FUNCTION_BLOCK basicMotorGenerico (* Logica unica do motor generico (partida direta ou inversor) *)
  (* Standard: 61499-2 *)
  (* Version 2.2, 12/11/2026, Hidryco, Hidryco, 2.2: cfgFalhaNA (contato de falha NA, dosagem 800). 2.1: raio do gerador vermelho (3) so com a carga liberada, a planta nos geradores E o motor ligado (igual ao Motor_VS, gradeamento e UV); liberado e parado = cinza (2). 2.0: velocidade da IHM/SCADA (stsVelocidadeIhm, antes stsVelocidadeHz) em %%: com inversor = fldVelocidadePct (LSP 0 %% a HSP 100 %%), sem inversor = 0 ou 100 %%; referencia e manual continuam em Hz. 1.9: velocidade manual (stpVelocidadeManual) em Hz; saidas stsVelocidadeHz/stsReferenciaHz para a IHM (conversao no CLP, 60 Hz = 100 %). 1.8: IHM: velocidade e referencia no maximo 1 vez por segundo com o motor ligado (antes a cada 0,1 %); o plug/processo (CNF_SPEED) continua na hora. 1.7: saida stsFalhaAtiva (falha presente agora: emergencia, termica, acionamento ou comunicacao) no CNF_HMI. 1.6: protecao termica nao memoriza - sai sozinha quando normaliza (sem reset). 1.5: reset so libera a falha de parada com o motor parado (antes liberava com o motor ainda ligado e a supervisao nao recomecava). 1.1: refeito no padrao SE.App2CommonProcess - eventos por grupo de dados, saidas so na mudanca, supervisao por E_DELAY (MON_T/MON_RESET/MON_MAX), horimetro e partidas pelo devMntCalc, escala linear com limites. 1.4: horimetro proprio com resolucao de 1 s (E_CYCLE + PERSISTENCE), termica NF por padrao *)
  PACKAGE Hidryco.HidrycoLib;
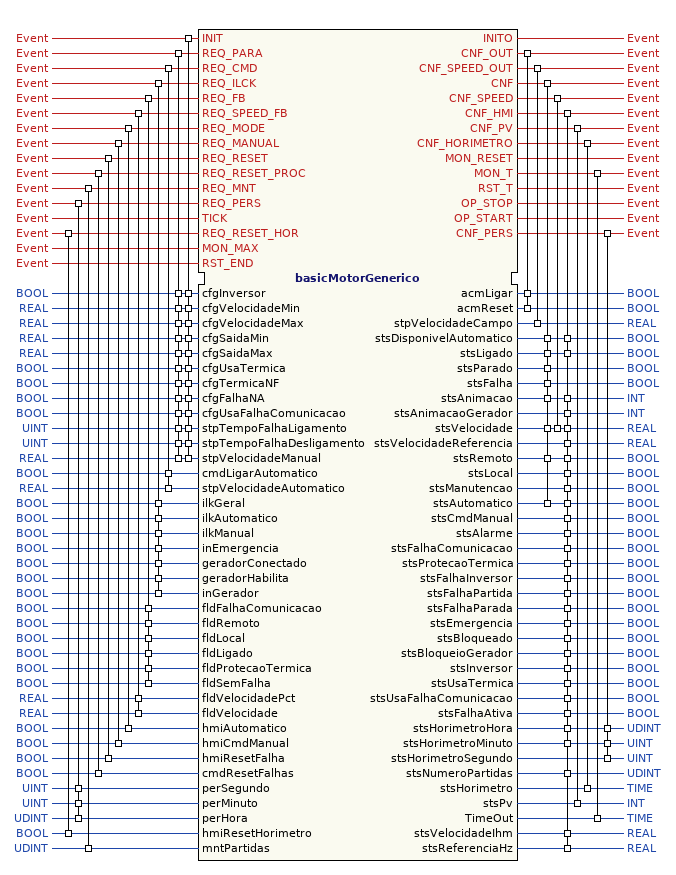
  EVENT_INPUT
    INIT WITH cfgInversor, cfgVelocidadeMin, cfgVelocidadeMax, cfgSaidaMin, cfgSaidaMax, cfgUsaTermica, cfgTermicaNF, cfgFalhaNA, cfgUsaFalhaComunicacao, stpTempoFalhaLigamento, stpTempoFalhaDesligamento, stpVelocidadeManual; (* Inicializacao (configuracao da instancia) *)
    REQ_PARA WITH cfgInversor, cfgVelocidadeMin, cfgVelocidadeMax, cfgSaidaMin, cfgSaidaMax, cfgUsaTermica, cfgTermicaNF, cfgFalhaNA, cfgUsaFalhaComunicacao, stpTempoFalhaLigamento, stpTempoFalhaDesligamento, stpVelocidadeManual; (* Atualizacao de parametros (IHM) *)
    REQ_CMD WITH cmdLigarAutomatico, stpVelocidadeAutomatico; (* Comando e referencia do processo *)
    REQ_ILCK WITH ilkGeral, ilkAutomatico, ilkManual, inEmergencia, geradorConectado, geradorHabilita, inGerador; (* Intertravamentos, emergencia e gerador *)
    REQ_FB WITH fldFalhaComunicacao, fldRemoto, fldLocal, fldLigado, fldProtecaoTermica, fldSemFalha; (* Sinais de campo *)
    REQ_SPEED_FB WITH fldVelocidade, fldVelocidadePct; (* Velocidade real do inversor *)
    REQ_MODE WITH hmiAutomatico; (* Modo automatico/manual (IHM) *)
    REQ_MANUAL WITH hmiCmdManual; (* Liga/desliga manual (IHM) *)
    REQ_RESET WITH hmiResetFalha; (* Reset de falhas (IHM) *)
    REQ_RESET_PROC WITH cmdResetFalhas; (* Reset de falhas (processo) *)
    REQ_MNT WITH mntPartidas; (* Numero de partidas do devMntCalc *)
    REQ_PERS WITH perSegundo, perMinuto, perHora; (* Horimetro lido do PERSISTENCE (READCNF) *)
    TICK; (* 1 s do E_CYCLE (so com o motor ligado) *)
    REQ_RESET_HOR WITH hmiResetHorimetro; (* Zera o horimetro (IHM) *)
    MON_MAX; (* Tempo de supervisao de partida/parada esgotado (E_DELAY) *)
    RST_END; (* Fim do pulso de reset (E_DELAY) *)
  END_EVENT
  EVENT_OUTPUT
    INITO; (* Inicializacao concluida *)
    CNF_OUT WITH acmLigar, acmReset; (* Saidas digitais de campo (na mudanca) *)
    CNF_SPEED_OUT WITH stpVelocidadeCampo; (* Referencia de velocidade para o campo (na mudanca) *)
    CNF WITH stsDisponivelAutomatico, stsLigado, stsParado, stsFalha, stsAnimacao, stsVelocidade, stsRemoto, stsAutomatico; (* Status para o processo (na mudanca) *)
    CNF_SPEED WITH stsVelocidade; (* Velocidade real (mudanca maior ou igual a 0,1 %) *)
    CNF_HMI WITH stsRemoto, stsLocal, stsManutencao, stsLigado, stsAutomatico, stsCmdManual, stsAnimacao, stsAnimacaoGerador, stsAlarme, stsFalhaComunicacao, stsProtecaoTermica, stsFalhaInversor, stsFalhaPartida, stsFalhaParada, stsEmergencia, stsBloqueado, stsBloqueioGerador, stsDisponivelAutomatico, stsVelocidade, stsVelocidadeReferencia, stsHorimetroHora, stsHorimetroMinuto, stsNumeroPartidas, stsInversor, stsUsaTermica, stsUsaFalhaComunicacao, stsFalhaAtiva, stsVelocidadeIhm, stsReferenciaHz; (* Status para a IHM (na mudanca) *)
    CNF_PV WITH stsPv; (* Estado ligado/parado para o devMntCalc (na mudanca) *)
    CNF_HORIMETRO WITH stsHorimetro; (* Tempo de operacao (na mudanca) *)
    MON_RESET; (* Cancela o tempo de supervisao (E_DELAY.STOP) - sai antes do MON_T *)
    MON_T WITH TimeOut; (* Inicia o tempo de supervisao (E_DELAY.START) *)
    RST_T; (* Inicia o pulso de reset (E_DELAY.START) *)
    OP_STOP; (* Para o E_CYCLE do horimetro - sai antes do OP_START *)
    OP_START; (* Inicia o E_CYCLE de 1 s do horimetro *)
    CNF_PERS WITH stsHorimetroSegundo, stsHorimetroMinuto, stsHorimetroHora; (* Grava o horimetro no PERSISTENCE (a cada minuto, na parada e no reset) *)
  END_EVENT
  VAR_INPUT
    cfgInversor : BOOL := FALSE; (* TRUE = motor com inversor (referencia de velocidade e medicoes) *)
    cfgVelocidadeMin : REAL := 0.0; (* Limite minimo da referencia de velocidade (%) *)
    cfgVelocidadeMax : REAL := 100.0; (* Limite maximo da referencia de velocidade (%) *)
    cfgSaidaMin : REAL := 0.0; (* Valor de campo equivalente a 0 % (referencia e realimentacao) *)
    cfgSaidaMax : REAL := 100.0; (* Valor de campo equivalente a 100 % (ex.: 100 = %, 60 = Hz, 10000 = Sulzer 0,01 %) *)
    cfgUsaTermica : BOOL := TRUE; (* TRUE = supervisiona a protecao termica *)
    cfgTermicaNF : BOOL := TRUE; (* TRUE = termica NF (FALSE no campo = atuada). Padrao NF (definido pelo usuario) *)
    cfgFalhaNA : BOOL := FALSE; (* TRUE = contato de falha do acionamento NA (TRUE no campo = falha, ligado em stsSemFalha). Padrao FALSE = NF (SEM FALHA) *)
    cfgUsaFalhaComunicacao : BOOL := TRUE; (* TRUE = considera o bit de falha de comunicacao da remota *)
    stpTempoFalhaLigamento : UINT; (* Tempo maximo para confirmar a partida (s). 0 = sem supervisao *)
    stpTempoFalhaDesligamento : UINT; (* Tempo maximo para confirmar a parada (s). 0 = sem supervisao *)
    stpVelocidadeManual : REAL; (* IHM: velocidade em manual em Hz (60 Hz = 100 %) *)
    cmdLigarAutomatico : BOOL; (* Comando ligar do processo (modo automatico) *)
    stpVelocidadeAutomatico : REAL; (* Referencia de velocidade do processo (%) *)
    ilkGeral : BOOL; (* Intertravamento geral (automatico e manual) *)
    ilkAutomatico : BOOL; (* Intertravamento so do automatico *)
    ilkManual : BOOL; (* Intertravamento so do manual *)
    inEmergencia : BOOL; (* Emergencia (TRUE = acionada): retira o comando e exige reset *)
    geradorConectado : BOOL; (* TRUE = o gerador pode alimentar este equipamento *)
    geradorHabilita : BOOL; (* Selecao do operador no CAT Gerador (HAB_GERADOR_EQUIP_n) *)
    inGerador : BOOL; (* TRUE = planta alimentada pelo gerador *)
    fldFalhaComunicacao : BOOL; (* Campo: falha de comunicacao da remota *)
    fldRemoto : BOOL; (* Campo: chave em remoto *)
    fldLocal : BOOL; (* Campo: chave em local *)
    fldLigado : BOOL; (* Campo: confirmacao de ligado *)
    fldProtecaoTermica : BOOL; (* Campo: protecao termica (ver cfgTermicaNF) *)
    fldSemFalha : BOOL; (* Campo: falha NF (TRUE = sem falha) *)
    fldVelocidadePct : REAL; (* Campo: velocidade do inversor em % (0 % no LSP, 100 % no HSP), so para a IHM *)
    fldVelocidade : REAL; (* Campo: velocidade real na unidade de cfgSaidaMin..cfgSaidaMax *)
    hmiAutomatico : BOOL; (* IHM: TRUE = automatico *)
    hmiCmdManual : BOOL; (* IHM: TRUE = ligar, FALSE = desligar (manual) *)
    hmiResetFalha : BOOL; (* IHM: reset de falhas (vale com TRUE) *)
    cmdResetFalhas : BOOL; (* Processo: reset de falhas (vale com TRUE) *)
    perSegundo : UINT; (* Horimetro persistido: segundos *)
    perMinuto : UINT; (* Horimetro persistido: minutos *)
    perHora : UDINT; (* Horimetro persistido: horas *)
    hmiResetHorimetro : BOOL; (* IHM: zera o horimetro (vale com TRUE) *)
    mntPartidas : UDINT; (* devMntCalc: numero de partidas *)
  END_VAR
  VAR_OUTPUT
    acmLigar : BOOL; (* Campo: comando liga *)
    acmReset : BOOL; (* Campo: pulso de reset (inversor/rele) *)
    stpVelocidadeCampo : REAL; (* Campo: referencia de velocidade (cfgSaidaMin..cfgSaidaMax) *)
    stsDisponivelAutomatico : BOOL; (* Pode ser comandado pelo automatico agora *)
    stsLigado : BOOL; (* Motor ligado (confirmacao de campo) *)
    stsParado : BOOL; (* Motor parado *)
    stsFalha : BOOL; (* Alguma falha memorizada (exige reset) *)
    stsAnimacao : INT; (* 0 desligado, 1 ligado, 2 falha, 3 manutencao *)
    stsAnimacaoGerador : INT; (* 0 nao conectado, 1 conectado, 2 selecionado, 3 selecionado e gerador ligado *)
    stsVelocidade : REAL; (* Velocidade real (%); partida direta: 0 ou 100 *)
    stsVelocidadeReferencia : REAL; (* Referencia de velocidade em uso (%) *)
    stsRemoto : BOOL; (* Chave em remoto *)
    stsLocal : BOOL; (* Chave em local *)
    stsManutencao : BOOL; (* Chave na posicao 0 *)
    stsAutomatico : BOOL; (* Modo automatico *)
    stsCmdManual : BOOL; (* Comando manual em vigor *)
    stsAlarme : BOOL; (* Falha memorizada ou falha de comunicacao *)
    stsFalhaComunicacao : BOOL; (* Falha de comunicacao *)
    stsProtecaoTermica : BOOL; (* Termica memorizada *)
    stsFalhaInversor : BOOL; (* Falha do acionamento memorizada *)
    stsFalhaPartida : BOOL; (* Nao confirmou partida no tempo *)
    stsFalhaParada : BOOL; (* Nao confirmou parada no tempo *)
    stsEmergencia : BOOL; (* Emergencia memorizada *)
    stsBloqueado : BOOL; (* Intertravamento ativo no modo atual *)
    stsBloqueioGerador : BOOL; (* Bloqueado pelo gerador *)
    stsInversor : BOOL; (* Copia de cfgInversor (IHM) *)
    stsUsaTermica : BOOL; (* Copia de cfgUsaTermica (IHM) *)
    stsUsaFalhaComunicacao : BOOL; (* Copia de cfgUsaFalhaComunicacao (IHM) *)
    stsFalhaAtiva : BOOL; (* Falha ativa (agora, sem memoria): emergencia, termica, acionamento ou comunicacao *)
    stsHorimetroHora : UDINT; (* Horimetro (h) *)
    stsHorimetroMinuto : UINT; (* Horimetro (min, 0-59) *)
    stsHorimetroSegundo : UINT; (* Horimetro (s, 0-59) *)
    stsNumeroPartidas : UDINT; (* Numero de partidas *)
    stsHorimetro : TIME; (* Tempo de operacao (IActStatus.FbHorimetro) *)
    stsPv : INT; (* Estado para o devMntCalc (0 parado, 1 ligado) *)
    TimeOut : TIME; (* Tempo de supervisao enviado ao E_DELAY *)
    stsVelocidadeIhm : REAL; (* Velocidade para a IHM/SCADA (%): com inversor entre LSP e HSP; sem inversor 0 ou 100 *)
    stsReferenciaHz : REAL; (* Referencia de velocidade em Hz (IHM/SCADA) *)
  END_VAR
  VAR
    initDone : BOOL; (* Bloco inicializado *)
    initPass : BOOL; (* Primeira execucao apos a inicializacao: envia tudo *)
    fbRecebido : BOOL; (* Ja recebeu a primeira leitura de campo *)
    bAutomatico : BOOL; (* Modo automatico (nao persistente) *)
    bCmdManual : BOOL; (* Comando manual memorizado (nao persistente) *)
    bComOk : BOOL; (* Comunicacao OK e campo ja lido *)
    bRemoto : BOOL;
    bLocal : BOOL;
    bLigado : BOOL;
    bManutencao : BOOL;
    bTermicaAtiva : BOOL; (* Termica atuada agora *)
    bFalhaInvAtiva : BOOL; (* Falha do acionamento presente agora *)
    bEmergencia : BOOL; (* Memoria de emergencia *)
    bTermica : BOOL; (* Memoria de termica *)
    bFalhaInversor : BOOL; (* Memoria de falha do acionamento *)
    bFalhaPartida : BOOL; (* Memoria de falha de partida *)
    bFalhaParada : BOOL; (* Memoria de falha de parada *)
    bFalha : BOOL; (* Alguma memoria de falha *)
    bReset : BOOL; (* Pedido de reset nesta execucao *)
    bResetPendente : BOOL; (* Pulso de reset em andamento *)
    bBloqueioGerador : BOOL;
    bPermissivo : BOOL; (* Pode operar (remoto, sem falha, sem bloqueio geral) *)
    iMon : INT; (* Supervisao: 0 nenhuma, 1 esperando ligar, 2 esperando desligar *)
    oldMon : INT; (* Supervisao em andamento no E_DELAY *)
    rRef : REAL; (* Referencia em % *)
    rFaixa : REAL; (* cfgSaidaMax - cfgSaidaMin *)
    wSts : WORD; (* Status da IHM em bits (deteccao de mudanca) *)
    oldSts : WORD := 16#FFFF;
    oldAcm : BOOL;
    oldReset : BOOL;
    oldStp : REAL := -1.0;
    oldStsProc : WORD := 16#FFFF;
    wStsProc : WORD; (* Status do processo em bits *)
    oldAnim : INT := -1;
    oldAnimGer : INT := -1;
    oldFalhaAtiva : BOOL;
    hmiRef : REAL := -1.0;
    hmiVel : REAL := -1.0;
    oldVel : REAL := -1.0;
    oldRef : REAL := -1.0;
    oldPv : INT := -1;
    oldHorimetro : TIME;
    oldMnt : UDINT := 16#FFFFFFFF;
    oldPartidas : UDINT := 16#FFFFFFFF;
    bPersLido : BOOL; (* Horimetro ja restaurado do PERSISTENCE *)
    bTick : BOOL; (* E_CYCLE do horimetro deve rodar *)
    oldTick : BOOL;
    uMinTotal : UDINT; (* Horimetro em minutos (deteccao de mudanca) *)
  END_VAR
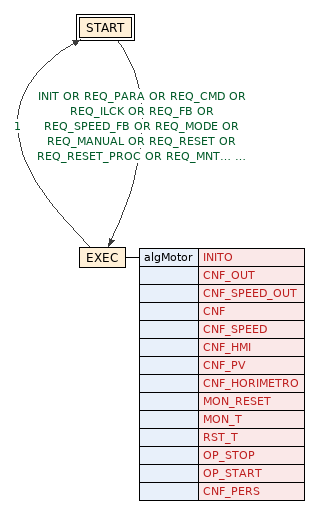
  EC_STATES
    START; (* Estado inicial *)
    EXEC : algMotor -> INITO, -> CNF_OUT, -> CNF_SPEED_OUT, -> CNF, -> CNF_SPEED, -> CNF_HMI, -> CNF_PV, -> CNF_HORIMETRO, -> MON_RESET, -> MON_T, -> RST_T, -> OP_STOP, -> OP_START, -> CNF_PERS; (* Executa a logica; o algoritmo decide quais eventos saem *)
  END_STATES
  EC_TRANSITIONS
    START TO EXEC := INIT OR REQ_PARA OR REQ_CMD OR REQ_ILCK OR REQ_FB OR REQ_SPEED_FB OR REQ_MODE OR REQ_MANUAL OR REQ_RESET OR REQ_RESET_PROC OR REQ_MNT OR REQ_PERS OR TICK OR REQ_RESET_HOR OR MON_MAX OR RST_END;
    EXEC TO START := 1;
  END_TRANSITIONS
  ALGORITHM algMotor IN ST: (* Logica completa do motor (um unico algoritmo) *)
(* =====================================================================
   basicMotorGenerico v1.1 - logica do CAT Motor_Generico (HidrycoLib)
   Padrao das bibliotecas Schneider (SE.App2CommonProcess):
   - eventos de saida desligados no inicio e ligados so na mudanca (variaveis oldX);
   - supervisao de partida/parada por E_DELAY externo (MON_T/MON_RESET/MON_MAX);
   - horimetro e partidas calculados e persistidos pelo devMntCalc.
   Regras de operacao (definidas pelo usuario):
   - emergencia, termica, falha do acionamento (NF), falha de partida e de
     parada ficam memorizadas ate o reset (IHM ou processo);
   - emergencia so retira o comando;
   - automatico -> manual mantem o motor como estava;
   - em manual o motor so liga com comando do operador: qualquer perda de
     permissivo cancela o comando manual (nao religa sozinho);
   - falha de comunicacao retira o comando, sem memorizar;
   - chave nem em local nem em remoto = manutencao.
   ===================================================================== *)

(* ---- 0. Eventos de saida: so sai o que for ligado abaixo ---- *)
INITO         := FALSE;
CNF_OUT       := FALSE;
CNF_SPEED_OUT := FALSE;
CNF           := FALSE;
CNF_SPEED     := FALSE;
CNF_HMI       := FALSE;
CNF_PV        := FALSE;
CNF_HORIMETRO := FALSE;
MON_RESET     := FALSE;
MON_T         := FALSE;
RST_T         := FALSE;
OP_STOP       := FALSE;
OP_START      := FALSE;
CNF_PERS      := FALSE;
bReset        := FALSE;

IF REQ_FB THEN
    fbRecebido := TRUE;                    (* campo valido a partir da 1a leitura *)
END_IF;

(* ---- 1. Inicializacao: nada e calculado antes do INIT ---- *)
IF INIT THEN
    initDone := TRUE;
    initPass := TRUE;
    INITO    := TRUE;
END_IF;
IF NOT initDone THEN
    RETURN;                                (* os dados recebidos ficam guardados *)
END_IF;

(* ---- 2. Sinais de campo (so atualizados com comunicacao OK) ---- *)
bComOk := fbRecebido AND NOT (cfgUsaFalhaComunicacao AND fldFalhaComunicacao);
IF bComOk THEN
    bRemoto := fldRemoto;
    bLocal  := fldLocal;
    bLigado := fldLigado;
    bTermicaAtiva  := cfgUsaTermica AND (fldProtecaoTermica XOR cfgTermicaNF);
    bFalhaInvAtiva := fldSemFalha XOR NOT cfgFalhaNA;   (* NF (padrao): FALSE no campo = falha; cfgFalhaNA: TRUE no campo = falha *)
ELSE
    bRemoto := FALSE;                      (* sem comunicacao: sai de remoto *)
    bLocal  := FALSE;
    bLigado := FALSE;                      (* e considera parado; memorias mantidas *)
END_IF;
bManutencao := bComOk AND NOT fldLocal AND NOT fldRemoto;

(* ---- 3. Falhas memorizadas ---- *)
IF inEmergencia THEN
    bEmergencia := TRUE;
END_IF;
IF bComOk THEN
    bTermica := bTermicaAtiva;             (* termica nao memoriza: sai sozinha quando normaliza *)
END_IF;
IF bComOk AND bFalhaInvAtiva THEN
    bFalhaInversor := TRUE;
END_IF;
(* tempo de supervisao esgotado: vale o tipo de espera que iniciou o E_DELAY *)
IF MON_MAX THEN
    IF oldMon = 1 THEN
        bFalhaPartida := TRUE;
    ELSIF oldMon = 2 THEN
        bFalhaParada := TRUE;
    END_IF;
END_IF;

(* ---- 4. Reset: libera so o que ja normalizou e pulsa o reset no campo ---- *)
bReset := (REQ_RESET AND hmiResetFalha) OR (REQ_RESET_PROC AND cmdResetFalhas);
IF bReset THEN
    IF NOT inEmergencia THEN
        bEmergencia := FALSE;
    END_IF;
    IF NOT bTermicaAtiva THEN
        bTermica := FALSE;
    END_IF;
    IF NOT bFalhaInvAtiva THEN
        bFalhaInversor := FALSE;
    END_IF;
    bFalhaPartida  := FALSE;
    IF NOT bLigado THEN
        bFalhaParada := FALSE;             (* so libera depois que o motor parou (sem comunicacao bLigado = FALSE) *)
    END_IF;
    bResetPendente := TRUE;
    RST_T          := TRUE;                (* pulso de reset para o campo *)
END_IF;
(* falha do acionamento que some durante o pulso de reset tambem e liberada *)
IF bResetPendente AND bComOk AND NOT bFalhaInvAtiva THEN
    bFalhaInversor := FALSE;
END_IF;
IF RST_END THEN
    bResetPendente := FALSE;
END_IF;
acmReset := bResetPendente;

(* ---- 5. Modo e comando manual (IHM) ---- *)
IF REQ_MODE THEN
    IF bAutomatico AND NOT hmiAutomatico THEN
        bCmdManual := acmLigar;            (* automatico -> manual: mantem como estava *)
    END_IF;
    bAutomatico := hmiAutomatico;
END_IF;
IF REQ_MANUAL THEN
    bCmdManual := hmiCmdManual;
END_IF;

(* ---- 6. Permissivos ---- *)
bFalha := bEmergencia OR bTermica OR bFalhaInversor OR bFalhaPartida OR bFalhaParada;
(* gerador: com a planta no gerador so opera o que esta conectado E selecionado *)
bBloqueioGerador := inGerador AND (NOT geradorConectado OR NOT geradorHabilita);
bPermissivo := bRemoto AND bComOk AND NOT bFalha AND NOT inEmergencia
               AND NOT bBloqueioGerador AND NOT ilkGeral;
IF NOT bPermissivo OR ilkManual THEN
    bCmdManual := FALSE;                   (* manual nunca religa sozinho *)
END_IF;

(* ---- 7. Comando ---- *)
acmLigar := bPermissivo AND
            ((bAutomatico AND cmdLigarAutomatico AND NOT ilkAutomatico) OR
             (NOT bAutomatico AND bCmdManual AND NOT ilkManual));

(* ---- 8. Supervisao de partida e parada (E_DELAY externo) ---- *)
IF bRemoto AND bComOk AND acmLigar AND NOT bLigado THEN
    iMon := 1;                             (* esperando confirmar ligado *)
ELSIF bRemoto AND bComOk AND NOT acmLigar AND bLigado THEN
    iMon := 2;                             (* esperando confirmar parado *)
ELSE
    iMon := 0;
END_IF;
IF iMon <> oldMon THEN
    MON_RESET := oldMon <> 0;              (* cancela a espera anterior *)
    IF iMon = 1 AND stpTempoFalhaLigamento > 0 THEN
        TimeOut := TO_TIME(UINT_TO_DINT(stpTempoFalhaLigamento) * 1000);
        MON_T := TRUE;
    ELSIF iMon = 2 AND stpTempoFalhaDesligamento > 0 THEN
        TimeOut := TO_TIME(UINT_TO_DINT(stpTempoFalhaDesligamento) * 1000);
        MON_T := TRUE;
    END_IF;
    oldMon := iMon;
END_IF;

(* ---- 9. Velocidade: limite em % e escala linear para o campo (como analogOutBasic) ---- *)
IF bAutomatico THEN
    rRef := stpVelocidadeAutomatico;
ELSE
    rRef := stpVelocidadeManual / 0.6;      (* IHM/SCADA em Hz (60 Hz = 100 %) -> % interno *)
END_IF;
IF cfgVelocidadeMax > cfgVelocidadeMin THEN
    rRef := LIMIT(cfgVelocidadeMin, rRef, cfgVelocidadeMax);
ELSE
    rRef := LIMIT(0.0, rRef, 100.0);
END_IF;
IF NOT cfgInversor THEN
    rRef := 0.0;                           (* partida direta: sem referencia *)
END_IF;
rFaixa := cfgSaidaMax - cfgSaidaMin;
IF rFaixa = 0.0 THEN
    rFaixa := 100.0;                       (* escala invalida: trata como % *)
END_IF;
stpVelocidadeCampo := cfgSaidaMin + rRef * rFaixa / 100.0;
IF cfgInversor THEN
    stsVelocidade := (fldVelocidade - cfgSaidaMin) * 100.0 / rFaixa;
ELSIF bLigado THEN
    stsVelocidade := 100.0;
ELSE
    stsVelocidade := 0.0;
END_IF;

(* ---- 10. Horimetro (resolucao de 1 s, persistido) e partidas (devMntCalc) ---- *)
(* sem comunicacao o estado fica congelado: evita contar partida falsa na volta *)
IF bComOk THEN
    IF bLigado THEN
        stsPv := 1;
    ELSE
        stsPv := 0;
    END_IF;
END_IF;
IF REQ_PERS THEN
    stsHorimetroSegundo := perSegundo;     (* restaura o valor gravado *)
    stsHorimetroMinuto  := perMinuto;
    stsHorimetroHora    := perHora;
    bPersLido := TRUE;
END_IF;
IF REQ_RESET_HOR AND hmiResetHorimetro THEN
    stsHorimetroSegundo := 0;
    stsHorimetroMinuto  := 0;
    stsHorimetroHora    := 0;
    CNF_PERS := TRUE;
END_IF;
IF TICK AND bTick THEN
    stsHorimetroSegundo := stsHorimetroSegundo + 1;
    IF stsHorimetroSegundo >= 60 THEN
        stsHorimetroSegundo := 0;
        stsHorimetroMinuto  := stsHorimetroMinuto + 1;
        CNF_PERS := TRUE;                  (* grava a cada minuto *)
        IF stsHorimetroMinuto >= 60 THEN
            stsHorimetroMinuto := 0;
            stsHorimetroHora   := stsHorimetroHora + 1;
        END_IF;
    END_IF;
END_IF;
(* E_CYCLE de 1 s so com o motor ligado; na parada grava os segundos acumulados *)
bTick := bPersLido AND (stsPv = 1);
IF bTick <> oldTick THEN
    IF bTick THEN
        OP_START := TRUE;
    ELSE
        OP_STOP  := TRUE;
        CNF_PERS := bPersLido;
    END_IF;
    oldTick := bTick;
END_IF;
uMinTotal := stsHorimetroHora * 60 + UINT_TO_UDINT(stsHorimetroMinuto);
stsNumeroPartidas := mntPartidas;
stsHorimetro := TO_TIME(UDINT_TO_LINT(stsHorimetroHora) * 3600000 + UINT_TO_LINT(stsHorimetroMinuto) * 60000 + UINT_TO_LINT(stsHorimetroSegundo) * 1000);

(* ---- 11. Status ---- *)
stsRemoto := bRemoto;
stsLocal := bLocal;
stsManutencao := bManutencao;
stsLigado := bLigado;
stsParado := NOT bLigado;
stsAutomatico := bAutomatico;
stsCmdManual := bCmdManual;
stsFalhaComunicacao := NOT bComOk;
stsProtecaoTermica := bTermica;
stsFalhaInversor := bFalhaInversor;
stsFalhaPartida := bFalhaPartida;
stsFalhaParada := bFalhaParada;
stsEmergencia := bEmergencia;
stsFalha := bFalha;
stsAlarme := bFalha OR NOT bComOk;
(* falha ativa (IHM STS_FALHA): condicao de falha presente agora, sem memoria nem reset *)
stsFalhaAtiva := inEmergencia OR NOT bComOk OR bTermicaAtiva OR bFalhaInvAtiva;
stsBloqueioGerador := bBloqueioGerador;
stsBloqueado := ilkGeral OR (bAutomatico AND ilkAutomatico) OR (NOT bAutomatico AND ilkManual);
stsDisponivelAutomatico := bAutomatico AND bPermissivo AND NOT ilkAutomatico;
stsVelocidadeReferencia := rRef;
(* velocidade para a IHM/SCADA em %: com inversor, leitura entre LSP (0 %) e HSP (100 %) do inversor *)
IF cfgInversor THEN
    stsVelocidadeIhm := fldVelocidadePct;
ELSE
    stsVelocidadeIhm := stsVelocidade;
END_IF;
stsReferenciaHz := rRef * 0.6;
(* configuracao para a IHM: os faceplates escondem o que nao se aplica ao tipo de motor *)
stsInversor := cfgInversor;
stsUsaTermica := cfgUsaTermica;
stsUsaFalhaComunicacao := cfgUsaFalhaComunicacao;

IF bManutencao THEN
    stsAnimacao := 3;
ELSIF bFalha THEN
    stsAnimacao := 2;
ELSIF bLigado THEN
    stsAnimacao := 1;
ELSE
    stsAnimacao := 0;
END_IF;

IF NOT geradorConectado THEN
    stsAnimacaoGerador := 0;
ELSIF NOT geradorHabilita THEN
    stsAnimacaoGerador := 1;
ELSIF inGerador AND bLigado THEN
    stsAnimacaoGerador := 3;              (* liberado, planta nos geradores e motor ligado *)
ELSE
    stsAnimacaoGerador := 2;              (* liberado, parado ou planta fora dos geradores *)
END_IF;

(* ---- 12. Emissao so na mudanca ---- *)
CNF_OUT := initPass OR (acmLigar <> oldAcm) OR (acmReset <> oldReset);
oldAcm := acmLigar;
oldReset := acmReset;

CNF_SPEED_OUT := initPass OR (stpVelocidadeCampo <> oldStp);
oldStp := stpVelocidadeCampo;

wStsProc := 16#0;
IF stsDisponivelAutomatico THEN wStsProc := wStsProc OR 16#0001; END_IF;
IF stsLigado THEN wStsProc := wStsProc OR 16#0002; END_IF;
IF stsFalha THEN wStsProc := wStsProc OR 16#0004; END_IF;
IF stsRemoto THEN wStsProc := wStsProc OR 16#0008; END_IF;
IF stsAutomatico THEN wStsProc := wStsProc OR 16#0010; END_IF;
CNF := initPass OR (wStsProc <> oldStsProc) OR (stsAnimacao <> oldAnim);
oldStsProc := wStsProc;

CNF_SPEED := initPass OR CNF OR (ABS(stsVelocidade - oldVel) >= 0.1);
IF CNF_SPEED THEN
    oldVel := stsVelocidade;
END_IF;

wSts := 16#0;
IF stsRemoto THEN wSts := wSts OR 16#0001; END_IF;
IF stsLocal THEN wSts := wSts OR 16#0002; END_IF;
IF stsManutencao THEN wSts := wSts OR 16#0004; END_IF;
IF stsLigado THEN wSts := wSts OR 16#0008; END_IF;
IF stsAutomatico THEN wSts := wSts OR 16#0010; END_IF;
IF stsCmdManual THEN wSts := wSts OR 16#0020; END_IF;
IF stsAlarme THEN wSts := wSts OR 16#0040; END_IF;
IF stsFalhaComunicacao THEN wSts := wSts OR 16#0080; END_IF;
IF stsProtecaoTermica THEN wSts := wSts OR 16#0100; END_IF;
IF stsFalhaInversor THEN wSts := wSts OR 16#0200; END_IF;
IF stsFalhaPartida THEN wSts := wSts OR 16#0400; END_IF;
IF stsFalhaParada THEN wSts := wSts OR 16#0800; END_IF;
IF stsEmergencia THEN wSts := wSts OR 16#1000; END_IF;
IF stsBloqueado THEN wSts := wSts OR 16#2000; END_IF;
IF stsBloqueioGerador THEN wSts := wSts OR 16#4000; END_IF;
IF stsDisponivelAutomatico THEN wSts := wSts OR 16#8000; END_IF;
CNF_HMI := initPass OR (wSts <> oldSts) OR (stsAnimacao <> oldAnim) OR (stsAnimacaoGerador <> oldAnimGer)
           OR (((TICK AND stsLigado) OR NOT stsLigado) AND ((stsVelocidade <> hmiVel) OR (rRef <> hmiRef)))   (* ligado: no maximo 1x/s *)
           OR (uMinTotal <> oldMnt) OR (mntPartidas <> oldPartidas)
           OR (stsFalhaAtiva <> oldFalhaAtiva);
oldFalhaAtiva := stsFalhaAtiva;
IF CNF_HMI THEN
    hmiVel := stsVelocidade; hmiRef := rRef;
END_IF;
oldSts := wSts;
oldAnim := stsAnimacao;
oldAnimGer := stsAnimacaoGerador;
oldRef := rRef;

CNF_PV := fbRecebido AND (stsPv <> oldPv);  (* so depois da 1a leitura do campo *)
oldPv := stsPv;

CNF_HORIMETRO := initPass OR (uMinTotal <> oldMnt);
oldMnt := uMinTotal;
oldPartidas := mntPartidas;

initPass := FALSE;
  END_ALGORITHM
END_FUNCTION_BLOCK
